TYPE "UDT_TestMotor"
VERSION : 0.1
   STRUCT
      Run : Bool := true;
      Speed : Real := 12.5;
      Total : DInt := 5000;
      Status : Word := 16#00A0;
      Descr : String[20] := 'motor';
   END_STRUCT;

END_TYPE
